Fanuc KAREL source: KT00830.KL

PROGRAM KT00830
%NOLOCKGROUP
VAR
  S1: STRING[80]
  S2: STRING[80]
  OUT: INTEGER
BEGIN
  S1 = 'A'
  S2 = 'B'
  S1 = 'A'
  S2 = 'B'
  OUT = SIN(S1)
END KT00830
